Fanuc KAREL source: KB00069.KL

PROGRAM KB00069
%NOLOCKGROUP
VAR
  P1: STRING[80]
  P2: INTEGER
  P3: STRING[80]
  P4: INTEGER
BEGIN
  P1 = 'A'
  P2 = 1
  P3 = 'A'
  P4 = 1
  DOSFILE_INF(P1, P2, P3, P4)
END KB00069
